(* IEC 61131-3 sources: Caravan/Archiv/12-04-19/Stations/MachineControl/MachineControl/Class/SafetyCDIAS_Base (part 4) *)

          // if it's our own path, remember the fast unsafe settings
          if (PathOfThisCPU[0]$UINT = (pListHeader^.p_us_Path$^UINT)^) & (To_StdLib.MemCmp(#PathOfThisCPU[0], pListHeader^.p_us_Path, PathOfThisCPU[0]$UINT + 2) = 0) then
            if (p_SDOResponseBuffer^.ud_Data <> 0) & (p_SDOResponseBuffer^.ud_Data <> 8) then
              b_FastUnsafeOutputsActive:= FALSE;

              // invalid number of fast unsafe output variables
              LogError("@ZZZZ (SafetyCDIAS_Base::ReadSDOConfig) Config Read Error: Invalid number of fast unsafe output vars (only 8 or 0 possible)");
            elsif (p_SDOResponseBuffer^.ud_Data = 8) then
              // if the client wasn't activated, we can't send anything
              if ActivateFastUnsafeIOs = 0 then
                b_FastUnsafeOutputsActive := FALSE;
                LogError("@ZZZZ (SafetyCDIAS_Base::ReadSDOConfig) Configuration Error: Fast unsafe outputs configured in safety designer but not activated at hardware class");
              else
                // otherwise we remember that we found the configuration and the client is set
                b_FastUnsafeOutputsActive := TRUE;
              end_if;
            else
              // no fast outputs configured via safety designer
              b_FastUnsafeOutputsActive := FALSE;
            end_if;
          end_if;
        end_if;

//*****************************************************************************
//**   UNSAFE BOOL OUTPUT VARIABLES                                          **
//*****************************************************************************

        //read number of unsafe output vars

        //send request and receive data
        sd_retval := SDOReadCfgRequ ( p_SDORequestBuffer  := p_SDORequestBuffer
                                    , p_SDOResponseBuffer := p_SDOResponseBuffer
                                    , ud_Address          := p_SDORequestBuffer^.ud_Address + 4
                                    , us_Length           := 4
                                    );

        //no response
        if ( sd_retval <> 0 ) then
          LogError("@ZZZZ (SafetyCDIAS_Base::ReadSDOConfig) Config Read Error: Reading number of unsafe bool output vars failed");
          return;
        end_if;

        ud_CntUnsafeOutputs := p_SDOResponseBuffer^.ud_Data;

        ud_Address := p_SDORequestBuffer^.ud_Address + 4;

        // skip the names of unsafe outputs
        for i := 1 to ud_CntUnsafeOutputs do

          // get length of Name
          sd_retval := SDOReadCfgRequ ( p_SDORequestBuffer  := p_SDORequestBuffer
                                      , p_SDOResponseBuffer := p_SDOResponseBuffer
                                      , ud_Address          := ud_Address
                                      , us_Length           := 4
                                      );
          //no response
          if ( sd_retval <> 0 ) then
            LogError("@ZZZZ (SafetyCDIAS_Base::ReadSDOConfig) Config Read Error: Reading length of unsafe bool output name failed");
            return;
          end_if;

          // prepare address to get name
          ud_Address    += 4;

          ud_TmpStrLen  := p_SDOResponseBuffer^.ud_Data;
          ud_ActStrLen  := ud_TmpStrLen;
          ud_TmpAddress := ud_Address;

          IF p_BlockedTransferMemory = NIL THEN
            sd_retval   := -100;
            ClassState  := _MemAllocFailed;
            RETURN;
          END_IF;

          IF ud_BlockedTransferMemorySize < (ud_TmpStrLen + 1) THEN
            p_BlockedTransferMemory := To_StdLib.ReAlloc(mptr:=p_BlockedTransferMemory, newsize:=(ud_TmpStrLen + 1));
            IF p_BlockedTransferMemory = NIL THEN
              ud_BlockedTransferMemorySize := 0;
              sd_retval   := -100;
              ClassState  := _MemAllocFailed;
              RETURN;
            ELSE
              ud_BlockedTransferMemorySize := (ud_TmpStrLen + 1);
            END_IF;
          END_IF;

          To_StdLib.MemSet(dest:=p_BlockedTransferMemory, value:=0, size:=ud_BlockedTransferMemorySize);

          p_TmpBlockedData := p_BlockedTransferMemory;

          us_BlockedTransferLength := BlockedTransferLength(ud_Datalength:=ud_TmpStrLen, us_MaxBlocklength:=60);

          while us_BlockedTransferLength do

            // get name
            sd_retval := SDOReadCfgRequ ( p_SDORequestBuffer  := p_SDORequestBuffer
                                        , p_SDOResponseBuffer := p_SDOResponseBuffer
                                        , ud_Address          := ud_TmpAddress
                                        , us_Length           := us_BlockedTransferLength
                                      );
            //no response
            if ( sd_retval <> 0 ) then
              LogError("@ZZZZ (SafetyCDIAS_Base::ReadSDOConfig) Config Read Error: Reading unsafe bool output name failed");
              return;
            end_if;

            To_StdLib.MemCpy(dest   := p_TmpBlockedData,
                             source := #p_SDOResponseBuffer^.ud_Data,
                             size   := us_BlockedTransferLength);

            p_TmpBlockedData  += us_BlockedTransferLength;
            ud_TmpAddress     += us_BlockedTransferLength;
            ud_TmpStrLen      -= us_BlockedTransferLength;

            us_BlockedTransferLength := BlockedTransferLength(ud_Datalength:=ud_TmpStrLen, us_MaxBlocklength:=60);

          end_while;

          sd_retval := AddUnsafeRoutElement(pRoutTable      := #p_UnsafeOutputsTable,
                                            pRoutElementsNo := #ui_CntUnsafeOutputs,
                                            ud_Address      := ud_ActAddress,
                                            ui_NameLen      := ud_ActStrLen$UINT,
                                            pNameNewElement := p_BlockedTransferMemory$^CHAR);

          // if unsafe component not found (sd_retval <> 0), it's not problem for whole safe application

          // get offset in application memory
          ud_ActAddress += 4;

          // prepare address for next unsafe output or for number of safe inputs
          ud_Address += ud_ActStrLen;

        end_for;

        // special unsafe variables (not supported by old modules)
        if b_CfgTypeV2 then

//*****************************************************************************
//**   UNSAFE BDINT OUTPUT VARIABLES                                         **
//*****************************************************************************

          //read number of unsafe BDINT output vars

          //send request and receive data
          sd_retval := SDOReadCfgRequ ( p_SDORequestBuffer  := p_SDORequestBuffer
                                      , p_SDOResponseBuffer := p_SDOResponseBuffer
                                      , ud_Address          := ud_Address
                                      , us_Length           := 4
                                      );

          //no response
          if ( sd_retval <> 0 ) then
            LogError("@ZZZZ (SafetyCDIAS_Base::ReadSDOConfig) Config Read Error: Reading number of unsafe BDINT output vars failed");
            return;
          end_if;

          ud_CntUnsafeOutputs := p_SDOResponseBuffer^.ud_Data;

          ud_Address := p_SDORequestBuffer^.ud_Address + 4;

          if ud_CntUnsafeOutputs then

            //SDO request for this command has 5 bytes additional data
            pBitMasks$^void := To_StdLib.Malloc(size := ud_CntUnsafeOutputs * sizeof(BDINT));

            if ( pBitMasks = NIL ) then
              sd_retval  := -100;
              ClassState := _MemAllocFailed;
              LogError("@ZZZZ (SafetyCDIAS_Base::ReadSDOConfig) Config Read Error: Failed to allocate memory for the BDINT variable bitmasks");
              return;
            end_if;

            // get the bitmasks for the BDINT variables
            for i := 1 to ud_CntUnsafeOutputs do

              // get bitmask
              sd_retval := SDOReadCfgRequ ( p_SDORequestBuffer  := p_SDORequestBuffer
                                          , p_SDOResponseBuffer := p_SDOResponseBuffer
                                          , ud_Address          := ud_Address
                                          , us_Length           := 4
                                          );
              //no response
              if ( sd_retval <> 0 ) then
                LogError("@ZZZZ (SafetyCDIAS_Base::ReadSDOConfig) Config Read Error: Reading bit mask of unsafe BDINT output failed");
                return;
              end_if;

              // prepare address for the next one
              ud_Address += 4;

              // save the bitmask for adding the rout element
              (pBitMasks + (i-1) * sizeof(BDINT))^ := p_SDOResponseBuffer^.ud_Data;
            end_for;

            // skip the names of unsafe outputs
            for i := 1 to ud_CntUnsafeOutputs do

              // get length of Name
              sd_retval := SDOReadCfgRequ ( p_SDORequestBuffer  := p_SDORequestBuffer
                                          , p_SDOResponseBuffer := p_SDOResponseBuffer
                                          , ud_Address          := ud_Address
                                          , us_Length           := 4
                                          );
              //no response
              if ( sd_retval <> 0 ) then
                LogError("@ZZZZ (SafetyCDIAS_Base::ReadSDOConfig) Config Read Error: Reading length of unsafe BDINT output name failed");
                return;
              end_if;

              // prepare address to get name
              ud_Address += 4;

              ud_TmpStrLen  := p_SDOResponseBuffer^.ud_Data;
              ud_ActStrLen  := ud_TmpStrLen;
              ud_TmpAddress := ud_Address;

              IF p_BlockedTransferMemory = NIL THEN
                sd_retval   := -100;
                ClassState  := _MemAllocFailed;
                RETURN;
              END_IF;

              IF ud_BlockedTransferMemorySize < (ud_TmpStrLen + 1) THEN
                p_BlockedTransferMemory := To_StdLib.ReAlloc(mptr:=p_BlockedTransferMemory, newsize:=(ud_TmpStrLen + 1));
                IF p_BlockedTransferMemory = NIL THEN
                  ud_BlockedTransferMemorySize := 0;
                  sd_retval := -100;
                  ClassState:= _MemAllocFailed;
                  RETURN;
                ELSE
                  ud_BlockedTransferMemorySize := (ud_TmpStrLen + 1);
                END_IF;
              END_IF;

              To_StdLib.MemSet(dest:=p_BlockedTransferMemory, value:=0, size:=ud_BlockedTransferMemorySize);

              p_TmpBlockedData := p_BlockedTransferMemory;

              us_BlockedTransferLength := BlockedTransferLength(ud_Datalength:=ud_TmpStrLen, us_MaxBlocklength:=60);

              while us_BlockedTransferLength do

                // get name
                sd_retval := SDOReadCfgRequ ( p_SDORequestBuffer  := p_SDORequestBuffer
                                            , p_SDOResponseBuffer := p_SDOResponseBuffer
                                            , ud_Address          := ud_TmpAddress
                                            , us_Length           := us_BlockedTransferLength
                                          );
                //no response
                if ( sd_retval <> 0 ) then
                  LogError("@ZZZZ (SafetyCDIAS_Base::ReadSDOConfig) Config Read Error: Reading unsafe BDINT output name failed");
                  return;
                end_if;

                To_StdLib.MemCpy(dest   := p_TmpBlockedData,
                                 source := #p_SDOResponseBuffer^.ud_Data,
                                 size   := us_BlockedTransferLength);

                p_TmpBlockedData          += us_BlockedTransferLength;
                ud_TmpAddress             += us_BlockedTransferLength;
                ud_TmpStrLen              -= us_BlockedTransferLength;

                us_BlockedTransferLength  := BlockedTransferLength(ud_Datalength:=ud_TmpStrLen, us_MaxBlocklength:=60);

              end_while;

              ActBitMask := (pBitMasks + (i-1) * sizeof(BDINT))^;

              sd_retval := AddUnsafeRoutElement(pRoutTable      := #p_UnsafeOutputsTable,
                                                pRoutElementsNo := #ui_CntUnsafeOutputs,
                                                ud_Address      := ud_UnsafeBDINT_Offset,
                                                ui_NameLen      := ud_ActStrLen$UINT,
                                                pNameNewElement := p_BlockedTransferMemory$^CHAR,
                                                BitMask         := ActBitMask);

              // if unsafe component not found (sd_retval <> 0), it's not problem for whole safe application

              // get offset in application memory
              ud_ActAddress         += CountBits(ActBitMask) * sizeof(DINT);
              ud_UnsafeBDINT_Offset += sizeof(DINT);

              // prepare address for next unsafe output or for number of safe inputs
              ud_Address            += ud_ActStrLen;

            end_for;

            // free the bitmasks
            To_StdLib.Free(mptr:=pBitMasks);
          end_if;
        end_if;

//*****************************************************************************
//**   SAFE INPUT VARIABLES                                                  **
//*****************************************************************************

        // get number of safe inputs
        sd_retval := SDOReadCfgRequ ( p_SDORequestBuffer  := p_SDORequestBuffer
                                    , p_SDOResponseBuffer := p_SDOResponseBuffer
                                    , ud_Address          := ud_Address
                                    , us_Length           := 4
                                    );

        //no response
        if ( sd_retval <> 0 ) then
          LogError("@ZZZZ (SafetyCDIAS_Base::ReadSDOConfig) Config Read Error: Reading number of safe inputs failed");
          return;
        end_if;

        //number of safe inputs
        ud_TmpCnt     := p_SDOResponseBuffer^.ud_Data;

        // get offset in application memory
        ud_ActAddress += ud_TmpCnt * 4;

        //address of path length of first safe input
        ud_Address    := p_SDORequestBuffer^.ud_Address + 4;

        //read path of all safe inputs and add them to routing lists
        for i := 1 to ud_TmpCnt do

          //read path
          sd_retval := ReadModulePath ( p_SDORequestBuffer          := p_SDORequestBuffer
                                      , p_SDOResponseBuffer         := p_SDOResponseBuffer
                                      , p_ud_Address                := #ud_Address
                                      , pModule                     := pModule
                                      , p_ud_ModulePathLen_Max      := #ud_ModulePathLen_Max
                                      , p_ud_ModulePathCompLen_Max  := #ud_ModulePathCompLen_Max
                                      , us_SDOMaxDataSize           := us_DataLength_Max
                                      );

          //no response, error
          if ( sd_retval <> 0 ) then
            LogError("@ZZZZ (SafetyCDIAS_Base::ReadSDOConfig) Config Read Error: Reading path of safe input failed");
            return;
          end_if;

          // if there is a valid module path
          if pModule^.p_us_Path <> NIL then
            //add module to routing tabs
            sd_retval := AddModuleToRoutingTabs ( pModule       := pModule
                                                , pListHeader   := pListHeader
                                                , b_IsOptional  := TempModuleConfig.Info.IsOptional
                                                );

            if (sd_retval <> 0 ) then
              if ( ClassState <> _ModFromCfgNotFound ) then
                LogError("@ZZZZ (SafetyCDIAS_Base::ReadSDOConfig) Config Read Error: Failed to add safe input module to routing tabs");
                return;
              end_if;
            end_if;
          end_if;

          //address of path length = last address + 2 * 4 bytes ( RemoteIndex + MaxAge)
          ud_Address += 8;

        end_for;

        if b_CfgTypeV3 then

//*****************************************************************************
//**   SAFE DINT INPUT VARIABLES                                             **
//*****************************************************************************

          // get number of safe DINT inputs
          sd_retval := SDOReadCfgRequ ( p_SDORequestBuffer  := p_SDORequestBuffer
                                      , p_SDOResponseBuffer := p_SDOResponseBuffer
                                      , ud_Address          := ud_Address
                                      , us_Length           := 4
                                      );

          //no response
          if ( sd_retval <> 0 ) then
            LogError("@ZZZZ (SafetyCDIAS_Base::ReadSDOConfig) Config Read Error: Reading number of safe DINT inputs failed");
            return;
          end_if;

          //number of safe inputs
          ud_TmpCnt     := p_SDOResponseBuffer^.ud_Data;

          // get offset in application memory
          ud_ActAddress += ud_TmpCnt * 4;

          //address of path length of first safe input
          ud_Address    := p_SDORequestBuffer^.ud_Address + 4;

          //read path of all safe inputs and add them to routing lists
          for i := 1 to ud_TmpCnt do

            //read path
            sd_retval := ReadModulePath ( p_SDORequestBuffer          := p_SDORequestBuffer
                                        , p_SDOResponseBuffer         := p_SDOResponseBuffer
                                        , p_ud_Address                := #ud_Address
                                        , pModule                     := pModule
                                        , p_ud_ModulePathLen_Max      := #ud_ModulePathLen_Max
                                        , p_ud_ModulePathCompLen_Max  := #ud_ModulePathCompLen_Max
                                        , us_SDOMaxDataSize           := us_DataLength_Max
                                        );

            //no response, error
            if ( sd_retval <> 0 ) then
              LogError("@ZZZZ (SafetyCDIAS_Base::ReadSDOConfig) Config Read Error: Reading path of safe DINT input failed");
              return;
            end_if;

            // if there is a valid module path
            if pModule^.p_us_Path <> NIL then
              //add module to routing tabs
              sd_retval := AddModuleToRoutingTabs ( pModule       := pModule
                                                  , pListHeader   := pListHeader
                                                  , b_IsOptional  := TempModuleConfig.Info.IsOptional
                                                  );

              if (sd_retval <> 0 ) then
                if ( ClassState <> _ModFromCfgNotFound ) then
                  LogError("@ZZZZ (SafetyCDIAS_Base::ReadSDOConfig) Config Read Error: Failed to add safe DINT input module to routing tabs");
                  return;
                end_if;
              end_if;
            end_if;

            //address of path length = last address + 2 * 4 bytes ( RemoteIndex + MaxAge)
            ud_Address += 8;

          end_for;
        end_if;

        // only available at new modules
        if b_CfgTypeV2 then

//*****************************************************************************
//**   SAFE INTERFACE INPUT VARIABLES                                        **
//*****************************************************************************

          // get number of safe interface input vars

          //send request and receive data
          sd_retval := SDOReadCfgRequ ( p_SDORequestBuffer  := p_SDORequestBuffer
                                      , p_SDOResponseBuffer := p_SDOResponseBuffer
                                      , ud_Address          := ud_Address
                                      , us_Length           := 4
                                      );

          //no response
          if ( sd_retval <> 0 ) then
            LogError("@ZZZZ (SafetyCDIAS_Base::ReadSDOConfig) Config Read Error: Reading number of safe interface input variables failed");
            return;
          end_if;

          // skip the number
          ud_Address += 4;

          //number of safe inputs
          ud_TmpCnt := p_SDOResponseBuffer^.ud_Data;

          // get offset in application memory
          ud_ActAddress += ud_TmpCnt * 4;

          if ud_TmpCnt then

            for i := 0 to (ud_TmpCnt-1) do
              // get length of the uncompressed path

              //send request and receive data
              sd_retval := SDOReadCfgRequ ( p_SDORequestBuffer  := p_SDORequestBuffer
                                          , p_SDOResponseBuffer := p_SDOResponseBuffer
                                          , ud_Address          := ud_Address
                                          , us_Length           := 4
                                          );

              //no response
              if ( sd_retval <> 0 ) then
                LogError("@ZZZZ (SafetyCDIAS_Base::ReadSDOConfig) Config Read Error: Reading length of uncompressed interface topology path failed");
                return;
              end_if;

              // skip length of top path
              ud_Address += 4;

              // skip top path
              ud_Address += p_SDOResponseBuffer^.ud_Data;

              // read length of compressed topology path

              //send request and receive data
              sd_retval := SDOReadCfgRequ ( p_SDORequestBuffer  := p_SDORequestBuffer
                                          , p_SDOResponseBuffer := p_SDOResponseBuffer
                                          , ud_Address          := ud_Address
                                          , us_Length           := 4
                                          );

              //no response
              if ( sd_retval <> 0 ) then
                LogError("@ZZZZ (SafetyCDIAS_Base::ReadSDOConfig) Config Read Error: Reading length of compressed interface topology path failed");
                return;
              end_if;

              // skip length of compressed top path
              ud_Address += 4;

              // skip compressed top path and remote index and maximum age
              ud_Address += p_SDOResponseBuffer^.ud_Data + 4 + 4;
            end_for;
          end_if;

(*
 4 Byte Anzahl
 4 Byte Länge vom Pfad, Pfad (vorne Pfad ":" dann CRC für da Interface dann bis auf 4 Byte aufgefüllt)
 4 Byte Länge vom komprimierten Pfad, komprimierter Pfad (vorne Pfad ":" dann CRC für da Interface dann bis auf 4 Byte aufgefüllt)
 4 Byte RemoteIndex
 4 Byte Maximales Alter
*)

        end_if;

        // only available at new containers
        if b_CfgTypeV3 then

//*****************************************************************************
//**   SAFE DINT INTERFACE INPUT VARIABLES                                   **
//*****************************************************************************

          // get number of safe DINT interface input vars

          //send request and receive data
          sd_retval := SDOReadCfgRequ ( p_SDORequestBuffer  := p_SDORequestBuffer
                                      , p_SDOResponseBuffer := p_SDOResponseBuffer
                                      , ud_Address          := ud_Address
                                      , us_Length           := 4
                                      );

          //no response
          if ( sd_retval <> 0 ) then
            LogError("@ZZZZ (SafetyCDIAS_Base::ReadSDOConfig) Config Read Error: Reading number of safe DINT interface input variables failed");
            return;
          end_if;

          // skip the number
          ud_Address += 4;

          //number of safe inputs
          ud_TmpCnt := p_SDOResponseBuffer^.ud_Data;

          // get offset in application memory
          ud_ActAddress += ud_TmpCnt * 4;

          if ud_TmpCnt then

            for i := 0 to (ud_TmpCnt-1) do
              // get length of the uncompressed path

              //send request and receive data
              sd_retval := SDOReadCfgRequ ( p_SDORequestBuffer  := p_SDORequestBuffer
                                          , p_SDOResponseBuffer := p_SDOResponseBuffer
                                          , ud_Address          := ud_Address
                                          , us_Length           := 4
                                          );

              //no response
              if ( sd_retval <> 0 ) then
                LogError("@ZZZZ (SafetyCDIAS_Base::ReadSDOConfig) Config Read Error: Reading length of uncompressed interface topology path failed at safe DINT input variables");
                return;
              end_if;

              // skip length of top path
              ud_Address += 4;

              // skip top path
              ud_Address += p_SDOResponseBuffer^.ud_Data;

              // read length of compressed topology path

              //send request and receive data
              sd_retval := SDOReadCfgRequ ( p_SDORequestBuffer  := p_SDORequestBuffer
                                          , p_SDOResponseBuffer := p_SDOResponseBuffer
                                          , ud_Address          := ud_Address
                                          , us_Length           := 4
                                          );

              //no response
              if ( sd_retval <> 0 ) then
                LogError("@ZZZZ (SafetyCDIAS_Base::ReadSDOConfig) Config Read Error: Reading length of compressed interface topology path failed at safe DINT input variables");
                return;
              end_if;

              // skip length of compressed top path
              ud_Address += 4;

              // skip compressed top path and remote index and maximum age
              ud_Address += p_SDOResponseBuffer^.ud_Data + 4 + 4;
            end_for;
          end_if;

(*
 4 Byte Anzahl
 4 Byte Länge vom Pfad, Pfad (vorne Pfad ":" dann CRC für da Interface dann bis auf 4 Byte aufgefüllt)
 4 Byte Länge vom komprimierten Pfad, komprimierter Pfad (vorne Pfad ":" dann CRC für da Interface dann bis auf 4 Byte aufgefüllt)
 4 Byte RemoteIndex
 4 Byte Maximales Alter
*)

        end_if;

//*****************************************************************************
//**   FAST UNSAFE INPUT VARIABLES                                           **
//*****************************************************************************

        // only available at new modules
        if b_CfgTypeV2 then

          // get number of fast unsafe intput vars (should be 8 or 0)

          //send request and receive data
          sd_retval := SDOReadCfgRequ ( p_SDORequestBuffer  := p_SDORequestBuffer
                                      , p_SDOResponseBuffer := p_SDOResponseBuffer
                                      , ud_Address          := ud_Address
                                      , us_Length           := 4
                                      );

          //no response
          if ( sd_retval <> 0 ) then
            LogError("@ZZZZ (SafetyCDIAS_Base::ReadSDOConfig) Config Read Error: Reading number of fast unsafe intput vars failed");
            return;
          end_if;

          ud_Address += 4;

          // get offset in application memory
          ud_ActAddress += p_SDOResponseBuffer^.ud_Data * 4;

          // if it's our own path, remember the fast unsafe settings
          if (PathOfThisCPU[0]$UINT = (pListHeader^.p_us_Path$^UINT)^) & (To_StdLib.MemCmp(#PathOfThisCPU[0], pListHeader^.p_us_Path, PathOfThisCPU[0]$UINT + 2) = 0) then
            if (p_SDOResponseBuffer^.ud_Data <> 0) & (p_SDOResponseBuffer^.ud_Data <> 8) then
              b_FastUnsafeInputsActive := FALSE;

              // invalid number of fast unsafe intput variables
              LogError("@ZZZZ (SafetyCDIAS_Base::ReadSDOConfig) Config Read Error: Invalid number of fast unsafe intput vars (only 8 or 0 possible)");
            elsif (p_SDOResponseBuffer^.ud_Data = 8) then
              // if the client wasn't activated, we can't send anything
              if ActivateFastUnsafeIOs = 0 then
                b_FastUnsafeInputsActive := FALSE;
                LogError("@ZZZZ (SafetyCDIAS_Base::ReadSDOConfig) Configuration Error: Fast unsafe inputs configured in safety designer but not activated at hardware class");
              else
                // otherwise we remember that we found the configuration and the client is set
                b_FastUnsafeInputsActive := TRUE;
              end_if;
            else
              // no fast inputs configured via safety designer
              b_FastUnsafeInputsActive := FALSE;

              if (b_FastUnsafeOutputsActive = FALSE) & ActivateFastUnsafeIOs then
                LogError("@ZZZZ (SafetyCDIAS_Base::ReadSDOConfig) Configuration Error: Fast unsafe outputs not configured in safety designer but activated at hardware class");
              end_if;
            end_if;
          end_if;
        end_if;

//*****************************************************************************
//**   UNSAFE BOOL INPUT VARIABLES                                           **
//*****************************************************************************

        // here we go for unsafe bool input vars

        // get number of unsafe input vars
        sd_retval := SDOReadCfgRequ ( p_SDORequestBuffer  := p_SDORequestBuffer
                                    , p_SDOResponseBuffer := p_SDOResponseBuffer
                                    , ud_Address          := ud_Address
                                    , us_Length           := 4
                                    );

        //no response
        if ( sd_retval <> 0 ) then
          LogError("@ZZZZ (SafetyCDIAS_Base::ReadSDOConfig) Config Read Error: Failed to read number of unsafe input vars");
          return;
        end_if;

        ud_CntUnsafeInputs := p_SDOResponseBuffer^.ud_Data;

        ud_Address := p_SDORequestBuffer^.ud_Address + 4;

        // skip the names of unsafe inputs
        for i := 1 to ud_CntUnsafeInputs do

          // get length of Name
          sd_retval := SDOReadCfgRequ ( p_SDORequestBuffer  := p_SDORequestBuffer
                                      , p_SDOResponseBuffer := p_SDOResponseBuffer
                                      , ud_Address          := ud_Address
                                      , us_Length           := 4
                                      );
          //no response
          if ( sd_retval <> 0 ) then
            LogError("@ZZZZ (SafetyCDIAS_Base::ReadSDOConfig) Config Read Error: Reading length of unsafe input name failed");
            return;
          end_if;

          // prepare address to get name
          ud_Address    += 4;

          ud_TmpStrLen  := p_SDOResponseBuffer^.ud_Data;
          ud_ActStrLen  := ud_TmpStrLen;
          ud_TmpAddress := ud_Address;

          IF p_BlockedTransferMemory = NIL THEN
            sd_retval   := -100;
            ClassState  := _MemAllocFailed;
            RETURN;
          END_IF;

          IF ud_BlockedTransferMemorySize < (ud_TmpStrLen + 1) THEN
            p_BlockedTransferMemory := To_StdLib.ReAlloc(mptr:=p_BlockedTransferMemory, newsize:=(ud_TmpStrLen + 1));
            IF p_BlockedTransferMemory = NIL THEN
              ud_BlockedTransferMemorySize  := 0;
              sd_retval                     := -100;
              ClassState                    := _MemAllocFailed;
              RETURN;
            ELSE
              ud_BlockedTransferMemorySize := (ud_TmpStrLen + 1);
            END_IF;
          END_IF;

          To_StdLib.MemSet(dest:=p_BlockedTransferMemory, value:=0, size:=ud_BlockedTransferMemorySize);

          p_TmpBlockedData          := p_BlockedTransferMemory;

          us_BlockedTransferLength  := BlockedTransferLength(ud_Datalength:=ud_TmpStrLen, us_MaxBlocklength:=60);

          while us_BlockedTransferLength do

          // get name
          sd_retval := SDOReadCfgRequ ( p_SDORequestBuffer  := p_SDORequestBuffer
                                      , p_SDOResponseBuffer := p_SDOResponseBuffer
                                      , ud_Address          := ud_TmpAddress
                                      , us_Length           := us_BlockedTransferLength
                                      );
          //no response
          if ( sd_retval <> 0 ) then
            LogError("@ZZZZ (SafetyCDIAS_Base::ReadSDOConfig) Config Read Error: Reading unsafe input name failed");
            return;
          end_if;

            To_StdLib.MemCpy(dest   := p_TmpBlockedData,
                             source := #p_SDOResponseBuffer^.ud_Data,
                             size   := us_BlockedTransferLength);

            p_TmpBlockedData += us_BlockedTransferLength;
            ud_TmpAddress += us_BlockedTransferLength;
            ud_TmpStrLen -= us_BlockedTransferLength;

            us_BlockedTransferLength := BlockedTransferLength(ud_Datalength:=ud_TmpStrLen, us_MaxBlocklength:=60);

          end_while;

          sd_retval := AddUnsafeRoutElement(pRoutTable      := #p_UnsafeInputsTable,
                                            pRoutElementsNo := #ui_CntUnsafeInputs,
                                            ud_Address      := ud_ActAddress,
                                            ui_NameLen      := ud_ActStrLen$UINT,
                                            pNameNewElement := p_BlockedTransferMemory$^CHAR);

          // if unsafe component not found (sd_retval <> 0), it's not problem for whole safe application

          // get offset in application memory
          ud_ActAddress += 4;

          // prepare address for next unsafe input
          ud_Address    += ud_ActStrLen;

        end_for;

        // only available at new modules
        if b_CfgTypeV2 then

//*****************************************************************************
//**   UNSAFE BDINT INPUT VARIABLES                                          **
//*****************************************************************************

          // here we go for unsafe BDINT input vars

          // get number of unsafe input vars
          sd_retval := SDOReadCfgRequ ( p_SDORequestBuffer  := p_SDORequestBuffer
                                      , p_SDOResponseBuffer := p_SDOResponseBuffer
                                      , ud_Address          := ud_Address
                                      , us_Length           := 4
                                      );

          //no response
          if ( sd_retval <> 0 ) then
            LogError("@ZZZZ (SafetyCDIAS_Base::ReadSDOConfig) Config Read Error: Failed to read number of unsafe BDINT input vars");
            return;
          end_if;

          ud_CntUnsafeInputs := p_SDOResponseBuffer^.ud_Data;

          ud_Address := p_SDORequestBuffer^.ud_Address + 4;

          if ud_CntUnsafeInputs then

            //SDO request for this command has 5 bytes additional data
            pBitMasks$^void := To_StdLib.Malloc(size := ud_CntUnsafeInputs * sizeof(BDINT));

            if ( pBitMasks = NIL ) then
              sd_retval                         := -100;
              ClassState := _MemAllocFailed;
              LogError("@ZZZZ (SafetyCDIAS_Base::ReadSDOConfig) Config Read Error: Failed to allocate memory for the BDINT variable bitmasks");
              return;
            end_if;

            // get the bitmasks for the BDINT variables
            for i := 1 to ud_CntUnsafeInputs do

              // get bitmask
              sd_retval := SDOReadCfgRequ ( p_SDORequestBuffer  := p_SDORequestBuffer
                                          , p_SDOResponseBuffer := p_SDOResponseBuffer
                                          , ud_Address          := ud_Address
                                          , us_Length           := 4
                                          );
              //no response
              if ( sd_retval <> 0 ) then
                LogError("@ZZZZ (SafetyCDIAS_Base::ReadSDOConfig) Config Read Error: Reading bit mask of unsafe BDINT input failed");
                return;
              end_if;

              // prepare address for the next one
              ud_Address += 4;

              // save the bitmask for adding the rout element
              (pBitMasks + (i-1) * sizeof(BDINT))^ := p_SDOResponseBuffer^.ud_Data;
            end_for;

            // get the names of unsafe inputs
            for i := 1 to ud_CntUnsafeInputs do

              // get length of Name
              sd_retval := SDOReadCfgRequ ( p_SDORequestBuffer  := p_SDORequestBuffer
                                          , p_SDOResponseBuffer := p_SDOResponseBuffer
                                          , ud_Address          := ud_Address
                                          , us_Length           := 4
                                          );
              //no response
              if ( sd_retval <> 0 ) then
                LogError("@ZZZZ (SafetyCDIAS_Base::ReadSDOConfig) Config Read Error: Reading length of unsafe BDINT input name failed");
                return;
              end_if;

              // prepare address to get name
              ud_Address += 4;

              ud_TmpStrLen := p_SDOResponseBuffer^.ud_Data;
              ud_ActStrLen := ud_TmpStrLen;
              ud_TmpAddress := ud_Address;

              IF p_BlockedTransferMemory = NIL THEN
                sd_retval := -100;
                ClassState := _MemAllocFailed;
                RETURN;
              END_IF;

              IF ud_BlockedTransferMemorySize < (ud_TmpStrLen + 1) THEN
                p_BlockedTransferMemory := To_StdLib.ReAlloc(mptr:=p_BlockedTransferMemory, newsize:=(ud_TmpStrLen + 1));
                IF p_BlockedTransferMemory = NIL THEN
                  ud_BlockedTransferMemorySize  := 0;
                  sd_retval                     := -100;
                  ClassState                    := _MemAllocFailed;
                  RETURN;
                ELSE
                  ud_BlockedTransferMemorySize := (ud_TmpStrLen + 1);
                END_IF;
              END_IF;

              To_StdLib.MemSet(dest:=p_BlockedTransferMemory, value:=0, size:=ud_BlockedTransferMemorySize);

              p_TmpBlockedData          := p_BlockedTransferMemory;

              us_BlockedTransferLength  := BlockedTransferLength(ud_Datalength:=ud_TmpStrLen, us_MaxBlocklength:=60);

              while us_BlockedTransferLength do

                // get name
                sd_retval := SDOReadCfgRequ ( p_SDORequestBuffer  := p_SDORequestBuffer
                                            , p_SDOResponseBuffer := p_SDOResponseBuffer
                                            , ud_Address          := ud_TmpAddress
                                            , us_Length           := us_BlockedTransferLength
                                          );
                //no response
                if ( sd_retval <> 0 ) then
                  LogError("@ZZZZ (SafetyCDIAS_Base::ReadSDOConfig) Config Read Error: Reading unsafe BDINT input name failed");
                  return;
                end_if;

                To_StdLib.MemCpy(dest   := p_TmpBlockedData,
                                 source := #p_SDOResponseBuffer^.ud_Data,
                                 size   := us_BlockedTransferLength);

                p_TmpBlockedData          += us_BlockedTransferLength;
                ud_TmpAddress             += us_BlockedTransferLength;
                ud_TmpStrLen              -= us_BlockedTransferLength;

                us_BlockedTransferLength  := BlockedTransferLength(ud_Datalength:=ud_TmpStrLen, us_MaxBlocklength:=60);

              end_while;

              ActBitMask := (pBitMasks + (i-1) * sizeof(BDINT))^;

              sd_retval := AddUnsafeRoutElement(pRoutTable      := #p_UnsafeInputsTable,
                                                pRoutElementsNo := #ui_CntUnsafeInputs,
                                                ud_Address      := ud_UnsafeBDINT_Offset,
                                                ui_NameLen      := ud_ActStrLen$UINT,
                                                pNameNewElement := p_BlockedTransferMemory$^CHAR,
                                                BitMask         := ActBitMask);

              // if unsafe component not found (sd_retval <> 0), it's not problem for whole safe application

              // get offset in application memory
              ud_ActAddress         += CountBits(ActBitMask) * sizeof(DINT);
              ud_UnsafeBDINT_Offset += sizeof(DINT);

              // prepare address for next unsafe output or for number of constants
              ud_Address += ud_ActStrLen;

            end_for;

            // free the bitmasks
            To_StdLib.Free(mptr:=pBitMasks);
          end_if;

//*****************************************************************************
//**   CONSTANTS                                                             **
//*****************************************************************************

          // constants

          //send request and receive data
          sd_retval := SDOReadCfgRequ ( p_SDORequestBuffer  := p_SDORequestBuffer
                                      , p_SDOResponseBuffer := p_SDOResponseBuffer
                                      , ud_Address          := ud_Address
                                      , us_Length           := 4
                                      );

          //no response
          if ( sd_retval <> 0 ) then
            LogError("@ZZZZ (SafetyCDIAS_Base::ReadSDOConfig) Config Read Error: Reading number of constants failed");
            return;
          end_if;

          // skip number of constants
          ud_Address += 4;

          // skip constants
          ud_Address += p_SDOResponseBuffer^.ud_Data * 4;

          if b_CfgTypeV3 then

//*****************************************************************************
//**   DINT CONSTANTS                                                        **
//*****************************************************************************

            // constants

            //send request and receive data
            sd_retval := SDOReadCfgRequ ( p_SDORequestBuffer  := p_SDORequestBuffer
                                        , p_SDOResponseBuffer := p_SDOResponseBuffer
                                        , ud_Address          := ud_Address
                                        , us_Length           := 4
                                        );

            //no response
            if ( sd_retval <> 0 ) then
              LogError("@ZZZZ (SafetyCDIAS_Base::ReadSDOConfig) Config Read Error: Reading number of DINT constants failed");
              return;
            end_if;

            // skip number of dint constants
            ud_Address += 4;

            // skip constants (8 byte per DINT constant)
            ud_Address += p_SDOResponseBuffer^.ud_Data * 8;

          end_if;

//*****************************************************************************
//**   LOCAL OUTPUTS                                                         **
//*****************************************************************************

          // local outputs
          //send request and receive data
          sd_retval := SDOReadCfgRequ ( p_SDORequestBuffer  := p_SDORequestBuffer
                                      , p_SDOResponseBuffer := p_SDOResponseBuffer
                                      , ud_Address          := ud_Address
                                      , us_Length           := 4
                                      );

          //no response
          if ( sd_retval <> 0 ) then
            LogError("@ZZZZ (SafetyCDIAS_Base::ReadSDOConfig) Config Read Error: Reading number of local outputs failed");
            return;
          end_if;

          // skip number of local outputs
          ud_Address += 4;

          // skip local outputs
          //++pr
          // only available at new modules
          if b_CfgTypeV2 then
            ud_Address += p_SDOResponseBuffer^.ud_Data * 8; // Used-Flag, Modulkennung(SDIAS)
          else
            ud_Address += p_SDOResponseBuffer^.ud_Data * 4; // Used-Flag
          end_if;

          if b_CfgTypeV3 then

//*****************************************************************************
//**   LOCAL DINT OUTPUTS                                                    **
//*****************************************************************************

            // local outputs
            //send request and receive data
            sd_retval := SDOReadCfgRequ ( p_SDORequestBuffer  := p_SDORequestBuffer
                                        , p_SDOResponseBuffer := p_SDOResponseBuffer
                                        , ud_Address          := ud_Address
                                        , us_Length           := 4
                                        );

            //no response
            if ( sd_retval <> 0 ) then
              LogError("@ZZZZ (SafetyCDIAS_Base::ReadSDOConfig) Config Read Error: Reading number of local outputs failed");
              return;
            end_if;

            // skip number of local outputs
            ud_Address += 4;

            // skip local outputs
            //++pr
            // only available at new modules
            if b_CfgTypeV2 then
              ud_Address += p_SDOResponseBuffer^.ud_Data * 8; // Used-Flag, Modulkennung(SDIAS)
            else
              ud_Address += p_SDOResponseBuffer^.ud_Data * 4; // Used-Flag
            end_if;

          end_if;

//*****************************************************************************
//**   SAFE BOOL INTERFACE OUTPUT VARIABLES                                  **
//*****************************************************************************

          // safe bool interface output vars
          //send request and receive data
          sd_retval := SDOReadCfgRequ ( p_SDORequestBuffer  := p_SDORequestBuffer
                                      , p_SDOResponseBuffer := p_SDOResponseBuffer
                                      , ud_Address          := ud_Address
                                      , us_Length           := 4
                                      );

          //no response
          if ( sd_retval <> 0 ) then
            LogError("@ZZZZ (SafetyCDIAS_Base::ReadSDOConfig) Config Read Error: Reading number of safe BOOL interface output variables failed");
            return;
          end_if;

          // skip safe BOOL interface output variables
          ud_Address += 4;

          // count the interface output variables
          BoolOuts := p_SDOResponseBuffer^.ud_Data;

//*****************************************************************************
//**   SAFE DINT INTERFACE OUTPUT VARIABLES                                  **
//*****************************************************************************

          // safe dint interface output vars
          //send request and receive data
          sd_retval := SDOReadCfgRequ ( p_SDORequestBuffer  := p_SDORequestBuffer
                                      , p_SDOResponseBuffer := p_SDOResponseBuffer
                                      , ud_Address          := ud_Address
                                      , us_Length           := 4
                                      );

          //no response
          if ( sd_retval <> 0 ) then
            LogError("@ZZZZ (SafetyCDIAS_Base::ReadSDOConfig) Config Read Error: Reading number of safe DINT interface output variables failed");
            return;
          end_if;

          // skip number of safe dint interface output vars
          ud_Address += 4;

          // count the interface output variables
          DintOuts := p_SDOResponseBuffer^.ud_Data;

          if b_CfgTypeV3 then

//*****************************************************************************
//**   DYNAMIC PARAMETERS (e.g. for SSI Module)                              **
//*****************************************************************************
(*
Version of Parameters is saved in hd_DynParaVersion
if it's 16#0001, then we read out the number of parameters which will follow
*)
          end_if;

          // if there are interface variables
          if BoolOuts | DintOuts then
            // calculate the length of the interface frame
            TempPdoConfig.PdoLen := CalcPDOLength(BoolOuts, DintOuts);

            TempPdoConfig.Info                := 0;
            TempPdoConfig.Info.IsInterfacePDO := TRUE;
            TempPdoConfig.Info.IsOptional     := (ud_ActBlockType = BLKTYPE_CFG_MODULE_OPTIONAL);

            // if it's a broadcast => mark it
            if (TempPath[0]$UINT = 2) & (TempPath[0]$HDINT = INTERFACE_FRAME_BROADCAST) then
              TempPdoConfig.Info.IFBroadCast  := TRUE;
            end_if;

            // this is the source of the interface frame
            TempPdoConfig.SourcePathLen := pListHeader^.p_us_Path^$UINT + 2;
            TempPdoConfig.pSourcePath   := pListHeader^.p_us_Path;

            // and the destination
            TempPdoConfig.DestPathLen   := TempPath[0]$UINT + 2;
            TempPdoConfig.pDestPath     := #TempPath[0];

            // add the interface PDO to the list
            AddPdoToCfg(TempPdoConfig);

            TempModuleConfig.Info.IsInterfaceSource := TRUE;
            TempModuleConfig.Info.IsInterfaceDest   := FALSE;
            TempModuleConfig.InterfaceCRC := TempPdoConfig.InterfaceCRC;
          else
            TempModuleConfig.Info.IsInterfaceSource := FALSE;
            TempModuleConfig.Info.IsInterfaceDest   := FALSE;
            TempModuleConfig.InterfaceCRC           := 0;
          end_if;
        else
          TempModuleConfig.Info.IsInterfaceSource   := FALSE;
          TempModuleConfig.Info.IsInterfaceDest     := FALSE;
          TempModuleConfig.InterfaceCRC             := 0;
        end_if;

        // if it's our own path, remember the safety number
        if (PathOfThisCPU[0]$UINT = (pListHeader^.p_us_Path$^UINT)^) & (To_StdLib.MemCmp(#PathOfThisCPU[0], pListHeader^.p_us_Path, PathOfThisCPU[0]$UINT + 2) = 0) then
          TempModuleConfig.SafetyNbr := SafetyNumber;
        else
          TempModuleConfig.SafetyNbr := 0;
        end_if;

        // only when there is a manager
        if pSafetyManagerThis then
          AddModuleToCfg(TempModuleConfig);
        end_if;

//**********************************************************************************************************************************************************
      BLKTYPE_OLD_MODE_FLAG: // flag fore FW to use old config-mode
        // we need the old TimeSync config-type
        NewConfigType := ConfigState_Old;

//**********************************************************************************************************************************************************
      BLKTYPE_CFG_XML: // configuration for uploading the project to the safetydesigner (network placement information, names of bits,...)
        // no useful information here for us

//**********************************************************************************************************************************************************
    else
      // skip it = do nothing
//      TRACE("Found unhandled Blocktype in configuration");
//**********************************************************************************************************************************************************
    end_case;

    ud_ListBaseAddress := ud_ListLength_Address + ud_ListLength;
  end_while;

  if ( ( sd_retval = 0 ) & ( ClassState = _ModFromCfgNotFound ) ) then
    sd_retval := -1;
  end_if;

END_FUNCTION

FUNCTION VIRTUAL SafetyCDIAS_Base::SDOReadCfgRequ
	VAR_INPUT
		p_SDORequestBuffer 	  : ^SDORequReadConfig;
		p_SDOResponseBuffer 	: ^SDORespReadConfig;
		ud_Address 	          : UDINT;
		us_Length 	          : USINT;
	END_VAR
	VAR_OUTPUT
		sd_retval 	          : DINT;
	END_VAR

  //sequence number
  p_SDORequestBuffer^.StdHeader.SeqNr := us_CntSequNr;

  //increase counter for sequence number
  if us_CntSequNr < 16#7F then
    us_CntSequNr += 1;
  else
    us_CntSequNr := 0;
  end_if;

  //address
  p_SDORequestBuffer^.ud_Address    := ud_Address;

  //length of expected data
  p_SDORequestBuffer^.us_Length     := us_Length;

  //calculate CRC (starting with length of data until the end of command)
  p_SDORequestBuffer^.StdHeader.CRC := 0;

  //send request
  sd_retval := SAFETY_iSendRequest( uiMaster    := 0
                                  , pucNode     := p_ObjectPath
                                  , uiInLength  := sizeof(SDORequReadConfig)
                                  , pucInput    := p_SDORequestBuffer$^USINT
                                  , uiOutLength := sizeof(SDORespReadConfig) - sizeof(SDORespReadConfig.ud_Data) + us_Length
                                  , pucOutput   := p_SDOResponseBuffer$^USINT
                                  );

  //no response
  if ( sd_retval <> 0 ) then
    LogError("@ZZZZ (SafetyCDIAS_Base::SDOReadCfgRequ) SAFETY_iSendRequest failed");

    // we remember to retry in a few seconds
    b_ReadConfigFailed := TRUE;
    return;
  end_if;

  //check sequence number to exclude a possible wrong response
  if ( p_SDORequestBuffer^.StdHeader.SeqNr <> p_SDOResponseBuffer^.StdHeader.SeqNr ) then
    // we remember to retry in a few seconds
    b_ReadConfigFailed := TRUE;
    //log not routable SDOs
    LogValue("@ZZZZ (SafetyCDIAS_Base::SDOReadCfgRequ) Invalid Sequence number in SDO Standard Response. Got {0} instead of expected {1}", to_udint(p_SDOResponseBuffer^.StdHeader.SeqNr), to_udint(p_SDORequestBuffer^.StdHeader.SeqNr));
    return;
  end_if;

  //check returncode of SDO
  if ( p_SDOResponseBuffer^.us_Returncode <> SDO_RETCODE_OK ) then
    //log not routable SDOs
    LogValue("@ZZZZ (SafetyCDIAS_Base::SDOReadCfgRequ) Safety module {0}: Retcode of SDO Standard Response was invalid. Retcode: {1}", SafetyNumber$UDINT, to_udint(p_SDOResponseBuffer^.us_Returncode));

//    // when reading fails because safety designer is writing at the same moment
//    if p_SDOResponseBuffer^.us_Returncode = SDO_MICROCTRL_DIFFER then
      // we remember to retry in a few seconds
      b_ReadConfigFailed := TRUE;
//    end_if;

    return;
  end_if;

  //check length of read data
  if ( p_SDOResponseBuffer^.us_Length = 0 ) then
    LogError("@ZZZZ (SafetyCDIAS_Base::SDOReadCfgRequ) Response length is 0");
    sd_retval := -104;
    return;
  end_if;

END_FUNCTION

FUNCTION VIRTUAL SafetyCDIAS_Base::GetRoutingData
	VAR_OUTPUT
		sd_retval 	            : DINT;
	END_VAR
	VAR
		p_SDORequestBuffer 	    : ^SDORequReadConfig;
		p_SDOResponseBuffer 	  : ^SDORespReadConfig;
    Module                  : PathInfoType;
    ListHeader              : PathInfoType;
    NotAvailableStr         : ARRAY [0..99] OF CHAR;
    Time1, Time2            : UDINT;
	END_VAR

  InitPathInfo(#Module);
  InitPathInfo(#ListHeader);

  //SDO request for this command has 5 bytes additional data
  p_SDORequestBuffer$^void := To_StdLib.Malloc(size := sizeof(SDORequReadConfig));

  if ( p_SDORequestBuffer = NIL ) then
    State.uiIO_Flags				          := 0;
		State.uiIO_Flags.PhysicAccessOff  := 1;
    sd_retval                         := -100;
    ClassState                        := _MemAllocFailed;
    return;
  end_if;

  //SDO response for this command can have maximum additional data
  p_SDOResponseBuffer$^void := To_StdLib.Malloc(size := SDO_MAX_LENGTH);

  if ( p_SDOResponseBuffer = NIL ) then

    To_StdLib.Free(mptr := p_SDORequestBuffer);

    State.uiIO_Flags				          := 0;
		State.uiIO_Flags.PhysicAccessOff  := 1;
    sd_retval                         := -100;
    ClassState                        := _MemAllocFailed;
    return;
  end_if;

  //alloc memory for path of input-safety-module
  Module.p_us_Path$^void := To_StdLib.Malloc(size := 5);

  if ( Module.p_us_Path = NIL ) then

    To_StdLib.Free(mptr := p_SDORequestBuffer);
    To_StdLib.Free(mptr := p_SDOResponseBuffer);

    State.uiIO_Flags				          := 0;
		State.uiIO_Flags.PhysicAccessOff  := 1;
    sd_retval                         := -100;
    ClassState                        := _MemAllocFailed;
    return;
  end_if;

  //alloc memory for compressed path of input-safety-module
  Module.p_us_PathComp$^void := To_StdLib.Malloc(size := 5);

  if ( Module.p_us_PathComp = NIL ) then

    To_StdLib.Free(mptr := p_SDORequestBuffer);
    To_StdLib.Free(mptr := p_SDOResponseBuffer);
    To_StdLib.Free(mptr := Module.p_us_Path);

    State.uiIO_Flags				          := 0;
		State.uiIO_Flags.PhysicAccessOff  := 1;
    sd_retval                         := -100;
    ClassState                        := _MemAllocFailed;
    return;
  end_if;

  //alloc memory for path in list header
  ListHeader.p_us_Path$^void := To_StdLib.Malloc(size := 5);

  if ( ListHeader.p_us_Path = NIL ) then

    To_StdLib.Free(mptr := p_SDORequestBuffer);
    To_StdLib.Free(mptr := p_SDOResponseBuffer);
    To_StdLib.Free(mptr := Module.p_us_Path);
    To_StdLib.Free(mptr := Module.p_us_PathComp);

    State.uiIO_Flags				          := 0;
		State.uiIO_Flags.PhysicAccessOff  := 1;
    sd_retval                         := -100;
    ClassState                        := _MemAllocFailed;
    return;
  end_if;

  //alloc memory for path in list header
  ListHeader.p_us_PathComp$^void := To_StdLib.Malloc(size := 5);

  if ( ListHeader.p_us_PathComp = NIL ) then

    To_StdLib.Free(mptr := p_SDORequestBuffer);
    To_StdLib.Free(mptr := p_SDOResponseBuffer);
    To_StdLib.Free(mptr := Module.p_us_Path);
    To_StdLib.Free(mptr := Module.p_us_PathComp);
    To_StdLib.Free(mptr := ListHeader.p_us_Path);

    State.uiIO_Flags				          := 0;
		State.uiIO_Flags.PhysicAccessOff  := 1;
    sd_retval                         := -100;
    ClassState                        := _MemAllocFailed;
    return;
  end_if;

  b_ReadConfigFailed := FALSE;

  // if there is a revision in the configuration this variable changes to TRUE
  b_GotNewRevision := FALSE;

Time1 := OS_READMICROSEC();
  //read config data via SDOs and add safety modules to routing lists
  sd_retval := ReadSDOConfig( p_SDORequestBuffer      := p_SDORequestBuffer
                            , p_SDOResponseBuffer     := p_SDOResponseBuffer
                            , pModule                 := #Module
                            , pListHeader             := #ListHeader
                            );
Time2 := OS_READMICROSEC();
ud_ConfigReadTime := Time2 - Time1;

  // if there is no revision in the configuration => clear it
  if (b_GotNewRevision = FALSE) then

    // free memory, if available
    if pPrjNameStr & pPrjRevStr then
      To_StdLib.Free(pPrjNameStr);
    end_if;

    // use local memory to show "not available"
    _strcpy(dest:=#NotAvailableStr[0], src:="<not available>");
    PrjNameMemLen := _strlen(src:=#NotAvailableStr[0]);
    PrjNameStrLen := PrjRevStrLen := PrjNameMemLen - 1;
    pPrjNameStr   := pPrjRevStr := #NotAvailableStr[0];

    // write the strings to the string objects
    ShowProjectRevision();

    // there is no memory, so reset the pointer and length informations
    pPrjNameStr   := NIL;
    pPrjRevStr    := NIL;

    PrjNameMemLen := 0;
    PrjNameStrLen := 0;
    PrjRevStrLen  := 0;
  end_if;

  // if reading failed, because designer is writing at the same time => we try again in a few seconds
  if b_ReadConfigFailed then

    // next time we check for the configured state of the cpu
    b_CheckConfigured   := TRUE;

    // check again in background
    ClassState          := _ReinitConfig;

    // and wait at least 3 secs
    ud_LastCheckConfig  := ops.tAbsolute;

  // error in configuration -> no work
  elsif ( sd_retval <> 0 ) & (ClassState <> _ReinitConfig) then
    State.uiIO_Flags                  := 0;

    if ClassState = _WaitForSynchronicity then
      ClassState := _UnknownCfgError;
    end_if;

    LogError("@ZZZZ (SafetyCDIAS_Base::GetRoutingData) Reading Safety Configuration failed!");
  else
    // if it's still invalid, moving is possible and none of the connected modules has any reason to deactivate it (otherwise it would be inactive)
    if (b_MoveCommandInputActive = _Invalid) & (b_SafetyOnLocalCDIAS = FALSE) then
      b_MoveCommandInputActive := _Active;
    end_if;

    // we start the data object for continous writing to the module after we know that there is an input for this module and the move command is active
    if b_MoveCommandInputActive = _Active then
      b_StartDOs := TRUE;

      WalkThroughPDOMoverList(pList := #pPDOMoverListInputs, _Active);
    else
      if b_VaranAvailable & (sd_VaranType = 1) then
        MasterConnect.ResetDO( p_data_object := p_HandlePDOWrite$^DINT, us_state := VARAN_DO_NO_RUN, ud_bytes := MaxLengthPDOWrite);
      end_if;
      // tell all modules which think we can communicate via pdo mover, that this is not the case any more
      // for all module which are configured as safety inputs for this module
      // delete list with modules where communication (input) with pdo mover is defined
      WalkThroughPDOMoverList(pList := #pPDOMoverListInputs, _Inactive);
    end_if;

    if pPDOMoverListInputs then
      CleanupPDOMoverList(pList := #pPDOMoverListInputs);
    end_if;

    // if it's still invalid, moving is possible and none of the connected modules has any reason to deactivate it (otherwise it would be inactive)
    if (b_MoveCommandOutputActive = _Invalid) & (b_SafetyOnLocalCDIAS = FALSE) then
      b_MoveCommandOutputActive := _Active;
    end_if;

    // we start the data object for continous writing to the module after we know that there is an input for this module and the move command is active
    if b_MoveCommandOutputActive = _Active then
      // if the mover is active we have to activate the data objects for continous run
      if sd_VaranType = 1 then
        if b_PayloadSupport = FALSE then
          //set right address of do
          MasterConnect.SetNewDOAddressRd( p_data := pPDOReadData$^DINT, ud_address:= ( ui_MyPlace + OFFSET_SPDO_DATA ) );
        end_if;

        MasterConnect.ResetDO( p_data_object := p_HandlePDORead$^DINT, us_state := VARAN_DO_CONT_RUN, ud_bytes := MaxLengthPDORead);
      end_if;
      WalkThroughPDOMoverList(pList := #pPDOMoverListInputs, _Active);//ZoePat 27.12.2012 14:31  PRÜFEN OB DAS RICHTIG IST!!??!! evtl. muss Outputs hier hin...
    else
      // tell all modules which think we can communicate via pdo mover, that this is not the case any more
      // for all module which are configured as safety outputs for this module
      // delete list with modules where communication (output) with pdo mover is defined
      WalkThroughPDOMoverList(pList := #pPDOMoverListOutputs, _Inactive);
    end_if;

    if pPDOMoverListOutputs then
      CleanupPDOMoverList(pList := #pPDOMoverListOutputs);
    end_if;

    // read config succeeded, check update cycle of unsafe variables
    CheckUnsafeUpdateCycle();

    // last thing to do is to start realtime and cyclic work (they do nothing in _ReinitConfig state
    if ud_UnsafeVarsNotFound then
      ClassState            := _UnsafeVarNotFound;
      ud_UnsafeVarsNotFound := 0;
    else
      if us_SetBusReadyState = SetBusReadyFinished then
        // we're already synchron from a former configuration phase
        ClassState          := _SafetyClassOK;
      else
        ClassState          := _WaitForSynchronicity;
      end_if;
    end_if;

    // check for interface frame destination modules and mark them
    GetDestinationCRCs();

    // if there is a safety manager create a configuration message and send it to the safety manager
    if pSafetyManagerThis then
      CreateAndSendCfg();
    end_if;
  end_if;

  // free temporary configuration lists if there were any
  FreeCfgLists();

  //free allocated buffers
  To_StdLib.Free(mptr := p_SDORequestBuffer);
  To_StdLib.Free(mptr := p_SDOResponseBuffer);
  To_StdLib.Free(mptr := Module.p_us_Path);
  To_StdLib.Free(mptr := Module.p_us_PathComp);

  // maybe the listheader pointers have been already freed by ReadModulePath
  if ListHeader.p_us_Path then
    To_StdLib.Free(mptr := ListHeader.p_us_Path);
  end_if;
  if ListHeader.p_us_PathComp then
    To_StdLib.Free(mptr := ListHeader.p_us_PathComp);
  end_if;

END_FUNCTION

FUNCTION VIRTUAL SafetyCDIAS_Base::ReadModulePath
	VAR_INPUT
		p_SDORequestBuffer 	        : ^SDORequReadConfig;
		p_SDOResponseBuffer 	      : ^SDORespReadConfig;
		p_ud_Address 	              : ^UDINT;
		pModule 	                  : ^PathInfoType;
		p_ud_ModulePathLen_Max 	    : ^UDINT;
		p_ud_ModulePathCompLen_Max 	: ^UDINT;
		us_SDOMaxDataSize 	        : USINT;
	END_VAR
	VAR_OUTPUT
		sd_retval 	                : DINT;
	END_VAR
  VAR
    ud_ModulePathLen_Act      : UDINT;
    p_ud_ModulePath_Act       : ^UDINT;
  END_VAR

  //read length of module path

  //send request and receive data
  sd_retval := SDOReadCfgRequ ( p_SDORequestBuffer  := p_SDORequestBuffer
                              , p_SDOResponseBuffer := p_SDOResponseBuffer
                              , ud_Address          := p_ud_Address^
                              , us_Length           := 4
                              );

  //no response
  if ( sd_retval <> 0 ) then
    LogError("@ZZZZ (SafetyCDIAS_Base::ReadModulePath) Failed to read length of module path");
    return;
  end_if;

  //length of module path
  ud_ModulePathLen_Act := p_SDOResponseBuffer^.ud_Data;

  //length is zero, check compressed path
  if ( ud_ModulePathLen_Act > 0 ) then

    //resize buffer for path, if it's too small
    if ( ud_ModulePathLen_Act > p_ud_ModulePathLen_Max^ ) then

      pModule^.p_us_Path$^void := To_StdLib.ReAlloc(mptr := pModule^.p_us_Path$^void, newsize := ud_ModulePathLen_Act);

      if ( pModule^.p_us_Path = NIL ) then

        State.uiIO_Flags				          := 0;
        State.uiIO_Flags.PhysicAccessOff  := 1;
        sd_retval                         := -100;
        ClassState                        := _MemAllocFailed;
        return;
      end_if;

      //increase max. path length
      p_ud_ModulePathLen_Max^ := ud_ModulePathLen_Act;

    end_if;

    //read path

    //address of first byte of path
    p_ud_Address^ += 4;

    //set pointer to first byte of target buffer
    p_ud_ModulePath_Act := ( pModule^.p_us_Path )$^UDINT;

    //read path block by block, if path is longer than max. length
    while ( ud_ModulePathLen_Act > us_SDOMaxDataSize ) do

      //send request and receive data
      sd_retval := SDOReadCfgRequ ( p_SDORequestBuffer  := p_SDORequestBuffer
                                  , p_SDOResponseBuffer := p_SDOResponseBuffer
                                  , ud_Address          := p_ud_Address^
                                  , us_Length           := us_SDOMaxDataSize
                                  );

      //no response
      if ( sd_retval <> 0 ) then
        LogError("@ZZZZ (SafetyCDIAS_Base::ReadModulePath) Failed to read block of module path");
        return;
      end_if;

      //copy part of path
      To_StdLib.MemCpy(dest := p_ud_ModulePath_Act , source := #p_SDOResponseBuffer^.ud_Data, size := us_SDOMaxDataSize);

      //rest of path to be read
      ud_ModulePathLen_Act -= us_SDOMaxDataSize;

      //address of next block
      p_ud_Address^ += us_SDOMaxDataSize;

      //set pointer to next free byte of target buffer
      p_ud_ModulePath_Act += us_SDOMaxDataSize;

    end_while;

    //read last bytes of path

    //send request and receive data
    sd_retval := SDOReadCfgRequ ( p_SDORequestBuffer  := p_SDORequestBuffer
                                , p_SDOResponseBuffer := p_SDOResponseBuffer
                                , ud_Address          := p_ud_Address^
                                , us_Length           := ud_ModulePathLen_Act$USINT
                                );

    //no response
    if ( sd_retval <> 0 ) then
      LogError("@ZZZZ (SafetyCDIAS_Base::ReadModulePath) Failed to read last bytes of module path");
      return;
    end_if;

    To_StdLib.MemCpy(dest := p_ud_ModulePath_Act, source := #p_SDOResponseBuffer^.ud_Data, size := ud_ModulePathLen_Act);

    //address of next byte after path
    //address of last block + length of last read block
    p_ud_Address^ += ud_ModulePathLen_Act;
  else

    if pModule^.p_us_Path <> NIL then
      To_StdLib.Free(mptr := pModule^.p_us_Path);
      pModule^.p_us_Path := NIL;
    end_if;

    //address of compressed path
    p_ud_Address^ += 4;
  end_if;

// ============================================================================================================================

  // compressed module path starts here

  // read length of module path

  // send request and receive data
  sd_retval := SDOReadCfgRequ ( p_SDORequestBuffer  := p_SDORequestBuffer
                              , p_SDOResponseBuffer := p_SDOResponseBuffer
                              , ud_Address          := p_ud_Address^
                              , us_Length           := 4
                              );

  //no response
  if ( sd_retval <> 0 ) then
    LogError("@ZZZZ (SafetyCDIAS_Base::ReadModulePath) Failed to read length of compressed module path");
    return;
  end_if;

  //length of module path
  ud_ModulePathLen_Act := p_SDOResponseBuffer^.ud_Data;

  pModule^.ui_PathCompLen := to_uint(ud_ModulePathLen_Act);

  //if length is zero, leave method
  if ( ud_ModulePathLen_Act = 0 ) then
    if pModule^.p_us_PathComp <> NIL then
      To_StdLib.Free(mptr := pModule^.p_us_PathComp);
      pModule^.p_us_PathComp := NIL;
    end_if;

    // address of CRC
    p_ud_Address^ += 4;

    return;
  end_if;

  //resize buffer for path, if it's too small
  if ( ud_ModulePathLen_Act > p_ud_ModulePathCompLen_Max^ ) then

    pModule^.p_us_PathComp$^void := To_StdLib.ReAlloc(mptr := pModule^.p_us_PathComp$^void, newsize := ud_ModulePathLen_Act);

    if ( pModule^.p_us_PathComp = NIL ) then

      State.uiIO_Flags				          := 0;
      State.uiIO_Flags.PhysicAccessOff  := 1;
      sd_retval                         := -100;
      ClassState                        := _MemAllocFailed;
      return;
    end_if;

    //increase max. path length
    p_ud_ModulePathCompLen_Max^ := ud_ModulePathLen_Act;

  end_if;

  //read path

  //address of first byte of path
  p_ud_Address^ += 4;

  //set pointer to first byte of target buffer
  p_ud_ModulePath_Act := pModule^.p_us_PathComp$^UDINT;

  //read path block by block, if path is longer than max. length
  while ( ud_ModulePathLen_Act > us_SDOMaxDataSize ) do

    //send request and receive data
    sd_retval := SDOReadCfgRequ ( p_SDORequestBuffer  := p_SDORequestBuffer
                                , p_SDOResponseBuffer := p_SDOResponseBuffer
                                , ud_Address          := p_ud_Address^
                                , us_Length           := us_SDOMaxDataSize
                                );

    //no response
    if ( sd_retval <> 0 ) then
      LogError("@ZZZZ (SafetyCDIAS_Base::ReadModulePath) Failed to read block of compressed module path");
      return;
    end_if;

    //copy part of path
    To_StdLib.MemCpy(dest := p_ud_ModulePath_Act , source := #p_SDOResponseBuffer^.ud_Data, size := us_SDOMaxDataSize);

    //rest of path to be read
    ud_ModulePathLen_Act -= us_SDOMaxDataSize;

    //address of next block
    p_ud_Address^ += us_SDOMaxDataSize;

    //set pointer to next free byte of target buffer
    p_ud_ModulePath_Act += us_SDOMaxDataSize;

  end_while;

  //read last bytes of path

  //send request and receive data
  sd_retval := SDOReadCfgRequ ( p_SDORequestBuffer  := p_SDORequestBuffer
                              , p_SDOResponseBuffer := p_SDOResponseBuffer
                              , ud_Address          := p_ud_Address^
                              , us_Length           := ud_ModulePathLen_Act$USINT
                              );

  //no response
  if ( sd_retval <> 0 ) then
    LogError("@ZZZZ (SafetyCDIAS_Base::ReadModulePath) Failed to read last bytes of compressed module path");
    return;
  end_if;

  To_StdLib.MemCpy(dest := p_ud_ModulePath_Act, source := #p_SDOResponseBuffer^.ud_Data, size := ud_ModulePathLen_Act);

  //address of next byte after path
  //address of last block + length of last read block
  p_ud_Address^ += ud_ModulePathLen_Act;

END_FUNCTION

FUNCTION VIRTUAL SafetyCDIAS_Base::AddModuleToRoutingTabs
	VAR_INPUT
		pModule 	                : ^PathInfoType;
		pListHeader 	            : ^PathInfoType;
    b_IsOptional              : BOOL;
	END_VAR
	VAR_OUTPUT
		sd_retval 	              : DINT;
	END_VAR
  VAR
    p_TargetObject            : pVirtualBase;
    p_SafetyBase              : pVirtualBase;
    ud_IO_SafeNumber          : HDINT;
    ud_PDO_Buffer             : UDINT;
    pMoveCommandInputActive   : ^PDOMoveState;
    pMoveCommandOutputActive  : ^PDOMoveState;
    ud_MoveSourceDOHandle     : UDINT;
    ud_MoveSourceAddr         : UDINT;
    ud_MoveSourceOffset       : UDINT;
    MyPara 	                  : CmdStruct;
    MyResult                  : results;
  END_VAR

  // if the cpu is connected via varan there is a chance to activate the Move Command (only if all inputs for the cpu are also connected via VARAN)
  if b_VaranAvailable & (b_SafetyOnLocalCDIAS = FALSE) then
    pMoveCommandInputActive   := #b_MoveCommandInputActive;
    pMoveCommandOutputActive  := #b_MoveCommandOutputActive;
  else
    pMoveCommandInputActive   := NIL;
    pMoveCommandOutputActive  := NIL;
  end_if;

  // initialize with invalid value
  ud_MoveSourceAddr := 0;

  sd_retval         := -1;

  //get this-pointer of object in network that is located with transfered path
  p_TargetObject    := ( MasterConnect.GetObjectThisp(p_us_ObjectPath := pModule^.p_us_Path) )$pVirtualBase;

  //this-pointer found
  if ( p_TargetObject ) then

    //add output module

    //If found this-pointer equals the own this-pointer, then the module has to be added to output-list.
    //This module (CPU) provides the safety input values for the output module (path in list-header).
    if ( p_TargetObject = this ) then

      //the output module is addressed by the ListHeaderPath
      //get this-pointer of object in network that is located with transfered path
      p_TargetObject := ( MasterConnect.GetObjectThisp(p_us_ObjectPath := pListHeader^.p_us_Path) )$pVirtualBase;

      //this-pointer found
      if ( p_TargetObject ) then

        MyPara.uiCmd := CMD_SM_GET_MODULE_TYPE;
        sd_retval$iprStates := p_TargetObject^.NewInst(#MyPara, #MyResult);

        //check if it's a safety module
        if ( MyResult.aData[0]$UDINT = SM_TYPE_SAFETY_MODULE ) then

          //object is based on SafetyBase
          p_SafetyBase    := ( p_TargetObject )$pVirtualBase;

          //get pointer on PDO output buffer
          ud_PDO_Buffer   := GetPointer2PDOBuffer();

          //configure safety output module and receive safety number
          //inform the output module about safety number and object path of the safe CPU
          MyPara.uiCmd    := CMD_SM_CONFIG_SAFETY_OUTPUT;
          MyPara.aPara[0] := SafetyNumber$DINT;
          MyPara.aPara[1] := this$DINT;
          MyPara.aPara[2] := (GetPointer2PDOBuffer())$DINT;
          MyPara.aPara[3] := pModule$DINT;
          MyPara.aPara[4] := pMoveCommandOutputActive$DINT;
          MyPara.aPara[5] := ud_LocalMoveSourceAddr$DINT;
          MyPara.aPara[6] := b_IsOptional;
          if sd_VaranType = 1 then
            MyPara.aPara[7] := p_HandlePDORead$DINT;
          else
            MyPara.aPara[7] := ud_HandlePDOReadMoverDO$DINT;
          end_if;

          MyPara.aPara[8]     := 0$DINT;

          sd_retval$iprStates := p_SafetyBase^.NewInst(#MyPara, #MyResult);

          ud_IO_SafeNumber    := MyResult.aData[0]$UDINT;

//          //configure safety output module and receive safety number
//          //inform the output module about safety number and object path of the safe CPU
//          ud_IO_SafeNumber := p_SafetyBase^.ConfigSafetyOutput  ( ud_SafeNrCPU    := SafetyNumber
//                                                                , ud_thisp        := this$UDINT
//                                                                , ud_p_PDOBuffer  := GetPointer2PDOBuffer()
//                                                                , pObject         := pModule
//                                                                , pMoveActive     := pMoveCommandOutputActive
//                                                                , ud_HandleSourceDO := p_HandlePDORead$UDINT  // LanSte 28.05.2013 Payload support
//                                                                , ud_MoveSourceAddr := ud_LocalMoveSourceAddr
//                                                                , ud_MoveSourceOffset:= 0 //LanSte 28.05.2013 Payload support
//                                                                , b_IsOptional := b_IsOptional
//                                                                );

          //output module successfully configured
          if ( ud_IO_SafeNumber <> 0 ) then

            // add thispointer to list of modules which are configured to communicate via pdo mover (output)
            if pMoveCommandOutputActive & (pMoveCommandOutputActive^ <> _Inactive) then
              AddToPDOMoverList(p_SafetyBase, #pPDOMoverListOutputs);
            end_if;

            //add module to routing table
            sd_retval := AddRoutingElement( ud_SafeNumber       := ud_IO_SafeNumber
                                          , ud_thisp            := p_SafetyBase$UDINT
                                          , pObject             := pListHeader
                                          );
          else
            sd_retval := 0; // could be an optional module
          end_if;
        else
          LogError("@ZZZZ (SafetyCDIAS_Base::AddModuleToRoutingTabs) Config Read Error: Output module: Trying to add a non-safety module to safety routing table");
          LogHWPath("HW-Path of Module: {0}", pListHeader^.p_us_Path);
        end_if;
      else
        LogError("@ZZZZ (SafetyCDIAS_Base::AddModuleToRoutingTabs) Config Read Error: Output module: No Object of HW-class found for module to be added to safety routing table");
        LogHWPath("HW-Path of Module: {0}", pListHeader^.p_us_Path);
      end_if;

    //add other cpu module

    elsif pModule = pListHeader then

      //the output module is addressed by the ListHeaderPath
      //get this-pointer of object in network that is located with transfered path
      p_TargetObject := ( MasterConnect.GetObjectThisp(p_us_ObjectPath := pListHeader^.p_us_Path) )$pVirtualBase;

      //this-pointer found
      if ( p_TargetObject ) then

        //check if it's a safety module
        MyPara.uiCmd := CMD_SM_GET_MODULE_TYPE;
        sd_retval$iprStates := p_TargetObject^.NewInst(#MyPara, #MyResult);

        if ( MyResult.aData[0]$UDINT = SM_TYPE_SAFETY_MODULE ) then

          //object is based on SafetyBase
          p_SafetyBase := ( p_TargetObject )$pVirtualBase;

          //get safety number
          MyPara.uiCmd := CMD_SM_CONFIG_SAFETY_CPU;

          sd_retval$iprStates := p_SafetyBase^.NewInst(#MyPara, #MyResult);

          ud_IO_SafeNumber := MyResult.aData[0]$UDINT;

//          ud_IO_SafeNumber := p_SafetyBase^.ConfigSafetyCpu();

          if ( ud_IO_SafeNumber <> 0 ) then

            //add module to routing table
            sd_retval := AddRoutingElement( ud_SafeNumber       := ud_IO_SafeNumber
                                          , ud_thisp            := p_SafetyBase$UDINT
                                          , pObject             := pListHeader
                                          );
          else
            LogError("@ZZZZ (SafetyCDIAS_Base::AddModuleToRoutingTabs) Config Read Error: CPU module: 0 is an invalid safety number");
            LogHWPath("HW-Path of Module: {0}", pListHeader^.p_us_Path);

            b_ReInitMarker := TRUE;
          end_if;
        else
          LogError("@ZZZZ (SafetyCDIAS_Base::AddModuleToRoutingTabs) Config Read Error: CPU module: Trying to add a non-safety module to safety routing table");
          LogHWPath("HW-Path of Module: {0}", pListHeader^.p_us_Path);
        end_if;
      else
        LogError("@ZZZZ (SafetyCDIAS_Base::AddModuleToRoutingTabs) Config Read Error: CPU module: No Object of HW-class found for module to be added to safety routing table");
        LogHWPath("HW-Path of Module: {0}", pListHeader^.p_us_Path);
      end_if;

    //add input module

    else
      //It's a safety input module, so it has to be added to safety input list.
      //check if found object represents a safety module
      MyPara.uiCmd := CMD_SM_GET_MODULE_TYPE;
      sd_retval$iprStates := p_TargetObject^.NewInst(#MyPara, #MyResult);
      if ( MyResult.aData[0]$UDINT = SM_TYPE_SAFETY_MODULE ) then

        //object is based on SafetyBase
        p_SafetyBase := p_TargetObject;

        //configure safety input module and receive pointer on PDO-Buffer and safety number
        MyPara.uiCmd    := CMD_SM_CONFIG_SAFETY_INPUT;
        MyPara.aPara[0] := SafetyNumber$DINT;
        MyPara.aPara[1] := this$DINT;
        MyPara.aPara[2] := (#ud_PDO_Buffer)$DINT;
        MyPara.aPara[3] := pMoveCommandInputActive$DINT;
        MyPara.aPara[4] := (#ud_MoveSourceAddr)$DINT;
        MyPara.aPara[5] := (#ud_MoveSourceDOHandle)$DINT;
        MyPara.aPara[6] := (#ud_MoveSourceOffset)$DINT;
        sd_retval$iprStates := p_SafetyBase^.NewInst(#MyPara, #MyResult);

        ud_IO_SafeNumber := MyResult.aData[0]$UDINT;

//      //configure safety input module and receive pointer on PDO-Buffer and safety number
//      ud_IO_SafeNumber := p_SafetyBase^.ConfigSafetyInput ( ud_SafeNrCPU          := SafetyNumber
//                                                          , ud_thisp              := this$UDINT
//                                                          , p_PDOBuffer           := #ud_PDO_Buffer
//                                                          , pMoveActive           := pMoveCommandInputActive
//                                                          , p_ud_HandleSourceDO   := #ud_MoveSourceDOHandle
//                                                          , p_ud_MoveSourceAddr   := #ud_MoveSourceAddr
//                                                          , p_ud_MoveSourceOffset := #ud_MoveSourceOffset
//                                                          );
        //input module successfully configured
        if ( ud_IO_SafeNumber <> 0 ) then
          // only if the configuration affects our cpu, we add something to our PDO input buffer
          p_TargetObject := ( MasterConnect.GetObjectThisp(p_us_ObjectPath := pListHeader^.p_us_Path) )$pVirtualBase;

          //this-pointer found
          if ( p_TargetObject = this ) then

            // add thispointer to list of modules which are configured to communicate via pdo mover (input)
            if pMoveCommandInputActive & (pMoveCommandInputActive^ <> _Inactive) then
              AddToPDOMoverList(p_SafetyBase, #pPDOMoverListInputs);
            end_if;

            //add pointer on PDO output buffer of input module to list of incoming PDOs
          //add pointer on PDO output buffer of input module to list of incoming PDOs
          sd_retval := AddPDOToInputBuffer( ud_p2Buffer         := ud_PDO_Buffer
                                          , ud_HandleSourceDO   := ud_MoveSourceDOHandle //LanSte 28.05.2013 Payload support
                                          , ud_MoveSourceAddr   := ud_MoveSourceAddr
                                          , ud_MoveSourceOffset := ud_MoveSourceOffset //LanSte 28.05.2013 Payload support
                                          , ud_SafetyNr         := ud_IO_SafeNumber
                                          , b_IsOptional        := b_IsOptional);          else
            sd_retval := 0;
          end_if;

          if ( sd_retval = 0 ) then

            //add module to routing table
            sd_retval := AddRoutingElement( ud_SafeNumber       := ud_IO_SafeNumber
                                          , ud_thisp            := p_SafetyBase$UDINT
                                          , pObject             := pModule
                                          );

          else
            LogError("@ZZZZ (SafetyCDIAS_Base::AddModuleToRoutingTabs) Config Read Error: Input module: Failed to add module to input buffer");
            LogHWPath("HW-Path of Module: {0}", pListHeader^.p_us_Path);
          end_if;
        else
          // module in configuration, which is not physically available but hw-class is placed
          sd_retval := 0; // could be an optional module
        end_if;
      else
        LogError("@ZZZZ (SafetyCDIAS_Base::AddModuleToRoutingTabs) Config Read Error: Input module: Trying to add a non-safety module to safety routing table");
        LogHWPath("HW-Path of Module: {0}", pModule^.p_us_Path);
      end_if;
    end_if;
  else
    // module in configuration, which is not physically available and no hw-class is placed
    LogError("@ZZZZ (SafetyCDIAS_Base::AddModuleToRoutingTabs) Config Read Error: Module in safety configuration, where no HW-Class is placed (maybe optional module)");
    LogHWPath("HW-Path of Module: {0}", pModule^.p_us_Path);
    sd_retval := 0;
  end_if;

END_FUNCTION

FUNCTION VIRTUAL SafetyCDIAS_Base::GetRoutingElementByThis
	VAR_INPUT
		ud_thisp 	        : UDINT;
	END_VAR
	VAR_OUTPUT
		p_RoutElement 	  : ^RoutElement;
	END_VAR
  VAR
  	i1                : UINT;
    p_RoutElement_Act : ^RoutElement;
  END_VAR

  p_RoutElement := NIL;

  //set pointer on first routing element
  p_RoutElement_Act := p_RoutTable;

  //check each element
  for i1 := 0 to ui_CntRoutElements - 1 do

    //if searched this is found, pointer on routing element is returned
    if ( p_RoutElement_Act^.ud_Thisp = ud_thisp ) then
      p_RoutElement := p_RoutElement_Act;
      return;
    end_if;

    //set pointer to next element
    p_RoutElement_Act += sizeof ( RoutElement );

  end_for;

END_FUNCTION

FUNCTION VIRTUAL SafetyCDIAS_Base::SDOStdRequ
	VAR_INPUT
		us_Command 	        : USINT;
		p_us_RespData 	    : ^USINT;
		us_RespLength 	    : USINT;
	END_VAR
	VAR_OUTPUT
		sd_retval 	        : DINT;
	END_VAR
  VAR
  	pSDORequestBuffer   : ^SDOStdHeader;
    pSDOResponseBuffer  : ^SDOStdResp;
    RespBuffer          : ARRAY [0..127] OF USINT;
    RequBuffer          : ARRAY [0..127] OF USINT;
    us_OutLength        : USINT;
  END_VAR

  //SDO requests for this commands don't have any further data
  pSDORequestBuffer$^void   := #RequBuffer[0];
  pSDOResponseBuffer$^void  := #RespBuffer[0];

  //SDO response buffer (length header + rc + data)
  us_OutLength := sizeof(SDOStdHeader) + 1 + us_RespLength;

  //calculate length without crc
  pSDORequestBuffer^.len    := sizeof(SDOStdHeader) - sizeof(SDOStdHeader.CRC);

  //type
  pSDORequestBuffer^.typ    := FRM_TYPECODE_STD;

  //sequence number
  pSDORequestBuffer^.SeqNr  := us_CntSequNr;

  //increase counter for sequence number
  if us_CntSequNr < 16#7F then
    us_CntSequNr += 1;
  else
    us_CntSequNr := 0;
  end_if;

  //command to inform CPU about initializing classes is ok
  pSDORequestBuffer^.cmd := us_Command;

  //set CRC-field to 0
  pSDORequestBuffer^.CRC := 0;

  //send request
  sd_retval := SAFETY_iSendRequest( uiMaster    := 0
                                  , pucNode     := p_ObjectPath
                                  , uiInLength  := sizeof(SDOStdHeader)
                                  , pucInput    := pSDORequestBuffer$^USINT
                                  , uiOutLength := us_OutLength
                                  , pucOutput   := pSDOResponseBuffer$^USINT
                                  );

  //no response
  if ( sd_retval = 0 ) then

    //check sequence number to exclude a possible wrong response
    if ( pSDORequestBuffer^.SeqNr <> pSDOResponseBuffer^.StdHeader.SeqNr ) then
      sd_retval := -102;
      //log not routable SDOs
      LogValue("@ZZZZ (SafetyCDIAS_Base::SDOStdRequ) Invalid Sequence number in SDO Standard Response. Got {0} instead of expected {1}", to_udint(pSDOResponseBuffer^.StdHeader.SeqNr), to_udint(pSDORequestBuffer^.SeqNr));

    //check returncode of SDO
    elsif ( pSDOResponseBuffer^.us_Returncode <> SDO_RETCODE_OK ) then
      //log not routable SDOs
      LogValue("@ZZZZ (SafetyCDIAS_Base::SDOStdRequ) Safety module {0}: Retcode of SDO Standard Response was invalid. Retcode: {1}", SafetyNumber$UDINT, to_udint(pSDOResponseBuffer^.us_Returncode));
      sd_retval := -103;
    end_if;
  else
    //log not routable SDOs
    LogValue("@ZZZZ (SafetyCDIAS_Base::SDOStdRequ) SAFETY_iSendRequest failed with retcode: -{0}", to_udint(ABS(sd_retval)));
  end_if;

  //return response
  if ( ( sd_retval = 0 ) & ( p_us_RespData <> NIL )) then

    To_StdLib.MemCpy(dest := p_us_RespData, source := #pSDOResponseBuffer^.us_Data, size := us_RespLength);

  end_if;

END_FUNCTION

FUNCTION VIRTUAL SafetyCDIAS_Base::GetPDOInputBuffer
	VAR_INPUT
		ud_p2Buffer 	    : UDINT;
	END_VAR
	VAR_OUTPUT
		p_InputBuffer 	  : ^PDOInputBuffer;
	END_VAR
  VAR
  	i1                : UINT;
    p_InputBuffer_Act : ^PDOInputBuffer;
  END_VAR

  p_InputBuffer := NIL;

  if ui_cnt_PDOInputBuffer then

    //set pointer on first input buffer element
    p_InputBuffer_Act := #aPDOInputBuffer[0];

    //check each element
    for i1 := 0 to (ui_cnt_PDOInputBuffer-1) do

      //if searched pointer is found, pointer on input buffer element is returned
      if ( p_InputBuffer_Act^.ud_p2Buffer = ud_p2Buffer ) then
        p_InputBuffer := p_InputBuffer_Act;
        return;
      end_if;

      //set pointer to next element
      p_InputBuffer_Act += sizeof ( PDOInputBuffer );

    end_for;
  end_if;

END_FUNCTION

FUNCTION VIRTUAL SafetyCDIAS_Base::GetThisViaServerName
	VAR_INPUT
		pObjectDotServer 	: ^CHAR;
	END_VAR
	VAR_OUTPUT
		ThisPtr 	        : pVoid;
	END_VAR
  VAR
    ChannelMode       : CHMODE;
  END_VAR

  ThisPtr := NIL;

  if pObjectDotServer = NIL then
    return;
  end_if;

  // get thispointer to server via name
  ChannelMode := _LookUpEmbed_C(pObjectDotServer, #ThisPtr, NIL);

  // check if it's a server
  case ChannelMode of
    _CH_CMD,
    _CH_SVR:

  else
    ThisPtr := NIL;
    LogError("@ZZZZ (SafetyCDIAS_Base::GetThisViaServerName) Couldn't get thispointer of server:");
    LogError(e_msg:=pObjectDotServer);
    ud_UnsafeVarsNotFound += 1;
  end_case;

END_FUNCTION

FUNCTION VIRTUAL SafetyCDIAS_Base::AddUnsafeRoutElement
	VAR_INPUT
		pRoutTable 	      : ^pUnsafeIORoutingElement;
		pRoutElementsNo 	: ^UINT;
		ud_Address 	      : UDINT;
		ui_NameLen 	      : UINT;
		pNameNewElement 	: ^CHAR;
		BitMask 	        : BDINT;
	END_VAR
	VAR_OUTPUT
		sd_retval 	      : DINT;
	END_VAR
  VAR
  	p_RoutElement     : ^UnsafeIORoutingElement;
    RemoteDomain      : USINT;
    LinearMemory      : BOOL;
  END_VAR

  sd_retval := -1;

  // check parameters
  if (ui_NameLen = 0) | (pNameNewElement = NIL) then
    LogError("@ZZZZ (SafetyCDIAS_Base::AddUnsafeRoutElement) Invalid call parameters for the variable name (invalid configuration in safety cpu)");
    return;
  end_if;

  // on CSCP011 the SDO_COMMAND_WRITE_VALUES didn't exist, so we have to make a difference here
  if (us_Variant = CSCP011_Preliminary) | (us_Variant = CSCP011_SERIES) | (pRoutTable = #p_UnsafeOutputsTable) then
    LinearMemory := TRUE;
  else
    LinearMemory := FALSE;
  end_if;

  // if there is a domain info attached
  if (pNameNewElement^ = '@') & ((pNameNewElement + 1)^ = 'D') then
    // check if it's in the actual domain
    if (pNameNewElement + 3)^ = ':' then
      // 1 digit domain number
      RemoteDomain := (pNameNewElement + 2)^ - '0';
    elsif (pNameNewElement + 4)^ = ':' then
      // 2 digits domain number
      RemoteDomain := ((pNameNewElement + 2)^ - '0') * 10 + (pNameNewElement + 3)^ - '0';
    else
      LogError("@ZZZZ (SafetyCDIAS_Base::AddUnsafeRoutElement) Invalid domain info at unsafe variable");
      return;
    end_if;

    // prepare the string (remove the domain info)
    if RemoteDomain >= 10 then
      ui_NameLen      -= 5;
      pNameNewElement += 5;
    else
      ui_NameLen      -= 4;
      pNameNewElement += 4;
    end_if;
  end_if;

  //With the first element, the table must be positioned
  if ( pRoutTable^ = NIL ) then

    //allocate memory for first routing element
    pRoutTable^$^void := To_StdLib.Malloc(size := sizeof(UnsafeIORoutingElement));

    if ( pRoutTable^ = NIL ) then

      State.uiIO_Flags                  := 0;
      State.uiIO_Flags.PhysicAccessOff 	:= 1;
      sd_retval                         :=-1;
      ClassState                        := _MemAllocFailed;
      return;

    end_if;

    p_RoutElement := pRoutTable^;

  else

    //add new element

    //add space for one element to table (linked list element for inputs and linear data area for outputs)
    if LinearMemory = FALSE then
    // search for a place
      p_RoutElement := pRoutTable^;
      while p_RoutElement^.pNext do
        p_RoutElement := p_RoutElement^.pNext;
      end_while;
      p_RoutElement^.pNext$^void := To_StdLib.Malloc(sizeof(UnsafeIORoutingElement));

      if ( p_RoutElement^.pNext = NIL ) then

        State.uiIO_Flags                  := 0;
        State.uiIO_Flags.PhysicAccessOff 	:= 1;
        sd_retval                         :=-1;
        ClassState                        := _MemAllocFailed;
        return;

      end_if;

      // set pointer to new element
      p_RoutElement := p_RoutElement^.pNext;
    else
      pRoutTable^$^void := To_StdLib.ReAlloc(mptr := pRoutTable^, newsize := ( ( pRoutElementsNo^ + 1 ) * sizeof(UnsafeIORoutingElement)));

      if ( pRoutTable^ = NIL ) then

        State.uiIO_Flags                  := 0;
        State.uiIO_Flags.PhysicAccessOff 	:= 1;
        sd_retval                         :=-1;
        ClassState                        := _MemAllocFailed;
        return;

      end_if;

      //set pointer to empty element on last position
      p_RoutElement := pRoutTable^ + ( pRoutElementsNo^ ) * sizeof(UnsafeIORoutingElement);
    end_if;
  end_if;

  if p_RoutElement then
    //allocate memory for name
    p_RoutElement^.pName$^void := To_StdLib.Malloc(size := ui_NameLen);
